FUNCTION_BLOCK FB_ForceController
(*

The function block used to 

Constructor: 		Patryk Panylo
Company:		E. Riexinger GmbH
Date:			17.02.2016
Version:			1.00

Date:			Revision:		Who:				Comment

*)
VAR_INPUT
	(* Input variables / Eingang Variablen *)
	bEnable					:BOOL;					(* Signal FB enable *)
	bControllerOn				:BOOL;					(* Controler on *)
	lrVeloKp					:LREAL := 0.1;				(* Kp Proportionalfaktor, deltaF x Kp -> v *)
	lrVeloTi					:LREAL := 10000;			(* Ti Integrationsfaktor*)
	lrCtrlVeloFilter				:LREAL := 0.01;			(* Control velocity filter =  0..1 *)
	lrPVForce				:LREAL;					(* Process variable of force *)
	lrSPForce				:LREAL;					(* Set point of force *)
	lrMaxForce				:LREAL;					(* Maximum force *)
	lrDeltaMax				:LREAL := 0.01;
	lrVeloMax				:LREAL := 10.0;			(* Maximum velocity [%] *)
	lrVeloMin				:LREAL := 0.0;				(* Minimum velocity [%] *)
	lrTaskCycle				:LREAL;					(* Task cycle *)
END_VAR
VAR_OUTPUT
	(* Output variables / Ausgang Variablen *)
	lrCVVelo					:LREAL;					(* Controller value of velocity [%] *)
END_VAR
VAR_IN_OUT
	(* Input Output variables / Ausgang Variablen *)

END_VAR
VAR
	(* Enummerations *)

	(* Variables *)

	(* References *)

	(* Interfaces *)

	(* Instances *)
	fbActForceFilter				:FB_ValueFilter;					(* Actual position filter *)
	fbCtrlPID						:FB_CtrlPID;

END_VAR
VAR CONSTANT

END_VAR


IF NOT bEnable
THEN
	lrCVVelo := 100;
	RETURN;
END_IF

(* Current force value filtering *)
fbActForceFilter(
	bEnable := TRUE,
	lrInSignal := lrPVForce,
	lrDeltaMax := lrDeltaMax,
);

IF bControllerOn
     AND fbActForceFilter.lrOutSignal < lrMaxForce
THEN

	fbCtrlPID(
		bEnable := TRUE,
		lrSetPoint := lrSPForce,
		lrProcessVariable := fbActForceFilter.lrOutSignal,
		lrDeadZone := 1.0,
		lrSignalOffset := 0.0,
		lrKp := lrVeloKp,
		lrTi := lrVeloTi,
		lrTd := 0.0,
		lrTaskCycle := lrTaskCycle,
		bManual := ,
		lrManualSignal:= ,
		lrLimitMin := lrVeloMin,
		lrLimitMax := lrVeloMax,
		lrProcessErr => ,
		bLimitMin => ,
		bLimitMax => );


	(*Reg_Rueck := Reg_Filt*Reg_Rueck + (1-Reg_Filt)*Reg_Verst*Drehzahl*Y_Vmax;*)
	(*lrCVVelo := MAX(0.0, (fbCtrlPID.lrCtrlVariable * (1.0 - lrPreCtrlVelo)) + (fbActForceFilter.lrOutSignal * lrPreCtrlVelo)); (* where lrPreCtrlVelo := 0.01 *)*)
	(*lrCVVelo := MAX(0.0, (fbCtrlPID.lrCtrlVariable * (1.0 - lrCtrlVeloFilter)) + (lrCVVelo * lrCtrlVeloFilter));				       (* where lrPreCtrlVelo := 0.99 *)*)
	lrCVVelo := MAX(0.0, (fbCtrlPID.lrCtrlVariable * lrCtrlVeloFilter) + (lrCVVelo * (1.0 - lrCtrlVeloFilter)));				       (* where lrPreCtrlVelo := 0.99 *)

ELSE
	lrCVVelo := 0.0;
END_IF

END_FUNCTION_BLOCK

(* stored: Version 1.1.0.1, ProductVersion 3.1.4024.15
   POU FB_ForceController: Id {72a41a0a-a576-4757-a8f0-fe478fddb194}, SpecialFunc None *)
